Staubli VAL3: bind.pgx

program bind()
  local string l_sbtn
  local num l_i
begin
  userPageBind("frame","lst1","options",sFrameList,size(sFrameList),"r")
  userPageBind("frame","lst2","options",sToolList,size(sToolList),"r")
  userPageBind("frame","lst1","value",sSelFrame,1,"rw")
  userPageBind("frame","lst2","value",sSelTool,1,"rw")
  //button
  for l_i =1 to 5
    l_sbtn="btn"+toString("",l_i)
    userPageBindClick("frame",l_sbtn,bBool[l_i],true)
  endFor
  userPageBindClick("frame","btnback",bBack,true)
end
